(* IEC 61131-3 sources: bcs-engineering-dsl/language/test/generating/after_test/expected, 2 files *)

(* ---- MAIN_decl.st ---- *)
PROGRAM MAIN
VAR
    conditionA: BOOL := TRUE;
    conditionB: BOOL := FALSE;
    AfterUnit_x: INT;
    TON_AfterInstance1: TON := (PT := T#5s);
    R_TRIG_AfterInstance1: R_TRIG;
    TON_AfterInstance2: TON := (PT := T#10s);
    R_TRIG_AfterInstance2: R_TRIG;
END_VAR

(* ---- MAIN_impl.st ---- *)
// Control Unit 'AfterUnit'
TON_AfterInstance1(IN := conditionA);
R_TRIG_AfterInstance1(CLK := TON_AfterInstance1.Q);
IF R_TRIG_AfterInstance1.Q THEN
    conditionB := TRUE;
    conditionA := FALSE;
END_IF;

TON_AfterInstance2(IN := conditionB = TRUE);
R_TRIG_AfterInstance2(CLK := TON_AfterInstance2.Q);
IF R_TRIG_AfterInstance2.Q THEN
    conditionA := TRUE;
    conditionB := FALSE;
END_IF;
